(* IEC 61131-3 sources: tsplc/packages/vscode-extension/tests/fixtures/conveyor/globals, 2 files *)

(* ---- PlantConstants.st ---- *)
{attribute 'qualified_only'}
VAR_GLOBAL CONSTANT
	ZoneCapacity : INT := 128;
END_VAR

(* ---- PlantIO.st ---- *)
{attribute 'qualified_only'}
VAR_GLOBAL
	Inbound : ST_Conveyor;
END_VAR
